(* IEC 61131-3 sources: ecmccfg/tests/integration/motion/ioc, 2 files *)

(* ---- motion.plc ---- *)
# Request/acknowledgement interface for manually driven acceptance cases.
# Capture each request once. Keep function return status separate from axis error.
VAR
  axis        : ax2;
  request     : static.request;
  ack         : static.ack;
  command     : static.command;
  target      : static.target;
  result      : static.result;
  commands    : static.commands;
  scans       : static.scans;
  firstScans  : static.firstScans;
  busy        : static.busy;
  homed       : static.homed;
  actual      : static.actual;
  enabled     : static.enabled;
  atTarget    : static.atTarget;
  axisError   : static.axisError;
  inputBit    : ec0.s3.binaryInput01;
  outputBit   : ec0.s4.binaryOutput01;
  ecValue     : static.ecValue;
  ecError     : static.ecError;
  dsError     : static.dsError;
  dsAverage   : static.dsAverage;
  encReady    : static.encReady;
  encHomed    : static.encHomed;
  hwReady     : static.hwReady;
  groupSize   : static.groupSize;
  groupMember : static.groupMember;
  groupBusy   : static.groupBusy;
  groupError  : static.groupError;
  groupEnable : static.groupEnable;
  seqRunning  : static.seqRunning;
  seqState    : static.seqState;
  lastTarget  : global.lastTarget;
  exchange    : global.exchange;
  exchangeAck : global.exchangeAck;
  peerAction  : global.peerAction;
  peerValue   : global.peerValue;
  privateVal  : static.privateVal;
  m2mPrevious : static.m2mPrevious;
END_VAR

if (${SELF}.firstscan) {
  firstScans := firstScans + 1;
};
scans := scans + 1;
var rc := 0;
if (request != ack) {
  if (command == 1) { rc := mc_power(2, 1); };
  if (command == 2) { rc := mc_power(2, 0); };
  if (command == 3) {
    mc_move_abs(2, 0, target, 0.15, 0.5, 0.5);
    if (abs(target) <= 0.6) {
      rc := mc_move_abs(2, 1, target, 0.15, 0.5, 0.5);
    } else { rc := -2; };
  };
  if (command == 4) {
    mc_move_rel(2, 0, target, 0.15, 0.5, 0.5);
    if (abs(mc_get_act_pos(2, 1) + target) <= 0.6) {
      rc := mc_move_rel(2, 1, target, 0.15, 0.5, 0.5);
    } else { rc := -2; };
  };
  if (command == 5) {
    mc_move_vel(2, 0, target, 0.5, 0.5);
    if (abs(target) <= 0.15) {
      rc := mc_move_vel(2, 1, target, 0.5, 0.5);
    } else { rc := -2; };
  };
  if (command == 6) { rc := mc_halt(2, 0); };
  if (command == 7) { rc := mc_reset(2); };
  if (command == 8) {
    mc_home_pos(2, 0, 15, 0.1, 0.1, 0);
    rc := mc_home_pos(2, 1, 15, 0.1, 0.1, 0);
  };
  if (command == 9) {
    ec_err_rst();
    var word := ec_set_bit(0, 3);
    word := ec_wrt_bit(word, 1, 0);
    word := ec_flp_bit(word, 1);
    word := ec_clr_bit(word, 0);
    word := ec_wrt_bits(word, 5, 4, 6);
    ecValue := word;
    outputBit := ec_chk_bit(word, 3) and ec_chk_bits(word, 4, 6) == 5 and inputBit;
    ec_set_bit(word, 64);
    ecError := ec_get_err();
    ec_err_rst();
    rc := ec_get_err();
  };
  if (command == 10) {
    ds_err_rst();
    rc := ds_clear_data(0) + ds_clear_data(1);
    if (ds_is_full(0) or ds_get_buff_id(0) != 0) { rc := -14; };
    rc := rc + ds_append_data(0, target);
    rc := rc + ds_append_data(0, target + 1);
    rc := rc + ds_append_data(0, target + 2);
    rc := rc + ds_append_data(0, target + 3);
    if (ds_get_size(0) != 4 or not(ds_is_full(0))) { rc := -10; };
    rc := rc + ds_set_buff_id(0, 2);
    if (ds_get_buff_id(0) != 2) { rc := -11; };
    rc := rc + ds_set_data(0, 2, target + 6);
    if (ds_get_data(0, 2) != target + 6) { rc := -12; };
    dsAverage := ds_get_avg(0);
    if (ds_get_min(0) != target or ds_get_max(0) != target + 6) { rc := -13; };
    rc := rc + ds_append_to_ds(0, 1, 2, 1);
    ds_append_to_ds(0, -1, 1, 1);
    dsError := ds_get_err();
    ds_err_rst();
    rc := rc + ds_get_err() + ds_push_asyn(0) + ds_push_asyn(1);
  };
  # 85000 = ERROR_MON_MAX_POSITION_LAG_EXCEEDED (0x14c08).
  if (command == 11) { rc := mc_set_axis_error(2, 85000); };
  if (command == 12) { rc := mc_grp_set_enable(0, target); };
  if (command == 13) { rc := mc_grp_halt(0); };
  if (command == 14) { rc := mc_grp_reset_error(0); };
  if (command == 15) {
    privateVal := target;
    peerValue := target;
    peerAction := 1;
    exchange := exchange + 1;
  };
  if (command == 16) { axis.traj.targetvel := target; };
  if (command == 17) {
    peerAction := target;
    exchange := exchange + 1;
  };
  if (command == 18) {
    m2m_err_rst();
    if (m2m_stat() != 1) {
      rc := m2m_get_err();
    } else {
      m2mPrevious := m2m_read(119);
      rc := m2m_write(119, target);
      if (rc == 0) {
        peerAction := 5;
        exchange := exchange + 1;
      };
    };
  };
  if (command == 19) { rc := m2m_write(119, m2mPrevious); };
  if (command == 20) { rc := mc_mr_set_stop(2, 1); };
  if (command == 21) {
    seq_arm(0, 0);
    rc := seq_arm(0, 1);
  };
  if (command < 1 or command > 21) { rc := -1; };
  result := rc;
  lastTarget := target;
  commands := commands + 1;
  ack := request;
};
busy := mc_get_busy(2);
homed := mc_get_homed(2);
actual := mc_get_act_pos(2, 1);
axisError := mc_get_axis_err(2);
enabled := axis.drv.enabled;
atTarget := axis.mon.attarget;
encReady := mc_get_enc_ready(2, 1);
encHomed := mc_get_enc_homed(2, 1);
hwReady := mc_get_hw_ready(2);
groupSize := mc_grp_size(0);
groupMember := mc_grp_axis_in_grp(0, 1) and mc_grp_axis_in_grp(0, 2);
groupBusy := mc_grp_get_any_busy(0);
groupError := mc_grp_get_any_error_id(0);
groupEnable := mc_grp_get_enabled(0);
seqRunning := seq_get_running(0);
seqState := seq_get_state(0);
static.axisId := axis.id;
static.axisPos := axis.enc.actpos;
static.axisTargetVel := axis.traj.targetvel;
static.seqValid := seq_get_valid(0);
static.seqArmed := seq_get_armed(0);

(* ---- peer.plc ---- *)
# Each request starts with one scan of writes. Read back on the next scan,
# after the PLC runtime has committed its direct data-interface writes.
VAR
  request : global.exchange;
  ack     : global.exchangeAck;
  action  : global.peerAction;
  value   : global.peerValue;
  localId : static.privateVal;
END_VAR

if (${SELF}.firstscan) { static.firstScans := static.firstScans + 1; };
static.scans := static.scans + 1;
static.scanTime := ${SELF}.scantime;
var scratch := 0;
scratch := scratch + 1;
static.localValue := scratch;

if (request != ack) {
  if (static.pending == 0) {
    if (action == 1) { localId := value + 100; };
    if (action == 2) { ds2.clear := 1; };
    if (action == 3) { ds2.append := localId; };
    if (action == 4) { ds2.index := 0; };
    if (action == 5) {
      static.m2mValue := m2m_read(119);
      static.m2mStatus := m2m_stat();
      m2m_read(-1);
      static.m2mError := m2m_get_err();
      m2m_err_rst();
      static.m2mErrorAfterReset := m2m_get_err();
    };
    if (action == 6) { ds2.data := localId + 1; };
    static.pending := 1;
  } else {
    static.storageSize := ds2.size;
    static.storageIndex := ds2.index;
    static.storageFull := ds2.full;
    static.storageData := ds2.data;
    static.storageError := ds2.error;
    ack := request;
    static.pending := 0;
  };
};
